(* IEC 61131-3 sources: SRCI_CLIENT_PLC/RobotLibrary/Library/POUs/Read/MC_ReadRobotData/Structures, 4 files *)

(* ---- ReadRobotDataOutCmd.st ---- *)
{attribute 'pack_mode' := '1'}
// -------------------------------------------------------------------------
//  SRCI Robot Library
// -------------------------------------------------------------------------
//
//  Object:      ReadRealsOutCmd
//  Author:      Thorsten Brach
//  Date:        2024-08-09
//
//  Description:
//
//
//  Copyright:
//    (C) 2024 Thorsten Brach. All rights reserved
//             Licensed under the MIT License.
//
//  Disclaimer:
//    This project is provided without any guarantee and can be used for
//    private and commercial purposes. Any use is at the user’s
//    own risk and responsibility.
//
// -------------------------------------------------------------------------
TYPE ReadRobotDataOutCmd :
STRUCT
  /// RC manufacturer name
  RCManufacturer       : STRING(20);
  /// RC part number
  RCOrderID            : STRING(20);
  /// RC serial number
  RCSerialNumber       : STRING(16);
  /// RA serial number
  RASerialNumber       : STRING(16);
  /// Robot firmware version in manufacturer -specific format
  RCFirmwareVersion    : STRING(12);
  ///
  /// Version of the server implementation in the format X.X.X (spec table 6-18) (ST-FIX F46: comment missing)
  RCInterpreterVersion : STRING(11); // ST-FIX F163: three numbers 0..255 as text 'M.m.p' (STRING(5) cut two-digit parts)
  /// Version of the SRCI interpreter on the RC as numbers (spec 6.1.2 table 6-11: Major, Minor, Patch) (ST-FIX F163: the text RCInterpreterVersion was decoded from single characters)
  RCInterpreterVersionNumber : VersionStruct;
  /// TRUE = Axis used in Robot FALSE = Axis NOT used. See Table 6-13 for bit assignment
  AxisJointUsed        : AxisJointUsed;
  /// TRUE = Axis used by Robot FALSE = Axis NOT used. See Table 6-13 for bit assignment.
  AxisExternalUsed     : AxisExternalUsed;
  /// TRUE = mm FALSE = ° See Table 6-13 for bit assignment.
  AxisJointUnit        : AxisJointUnit;
  /// TRUE = mm FALSE = ° See Table 6-13 for bit assignment
  AxisExternalUnit     : AxisExternalUnit;
  /// • TRUE: Function is supported by RC • FALSE: Function is not supported by RC See Table 6-14 for bit assignment.
  RCSupportedFunctions  : RCSupportedFunctions;
  /// Unique and unmodifiable identification of the RA.
  RobotID              : STRING(16);
  /// Interpreter task cycle time of the RC [ms]
  InterpreterCycleTime : UINT;
END_STRUCT
END_TYPE

(* ---- ReadRobotDataParCmd.st ---- *)
{attribute 'pack_mode' := '1'}
// -------------------------------------------------------------------------
//  SRCI Robot Library
// -------------------------------------------------------------------------
//
//  Object:      ReadRealsParCmd
//  Author:      Thorsten Brach
//  Date:        2024-08-09
//
//  Description:
//
//
//  Copyright:
//    (C) 2024 Thorsten Brach. All rights reserved
//             Licensed under the MIT License.
//
//  Disclaimer:
//    This project is provided without any guarantee and can be used for
//    private and commercial purposes. Any use is at the user’s
//    own risk and responsibility.
//
// -------------------------------------------------------------------------
TYPE ReadRobotDataParCmd :
STRUCT
END_STRUCT
END_TYPE

(* ---- ReadRobotDataRecvData.st ---- *)
{attribute 'pack_mode' := '1'}
// -------------------------------------------------------------------------
//  SRCI Robot Library
// -------------------------------------------------------------------------
//
//  Object:      ReadRealsRecvData
//  Author:      Thorsten Brach
//  Date:        2024-08-09
//
//  Description:
//
//
//  Copyright:
//    (C) 2024 Thorsten Brach. All rights reserved
//             Licensed under the MIT License.
//
//  Disclaimer:
//    This project is provided without any guarantee and can be used for
//    private and commercial purposes. Any use is at the user’s
//    own risk and responsibility.
//
// -------------------------------------------------------------------------
TYPE ReadRobotDataRecvData EXTENDS RspHeader :
STRUCT
  /// RC manufacturer name
  RCManufacturer       : STRING(20);
  /// RC part number
  RCOrderID            : STRING(20);
  /// RC serial number
  RCSerialNumber       : STRING(16);
  /// RA serial number
  RASerialNumber       : STRING(16);
  /// Robot firmware version in manufacturer -specific format
  RCFirmwareVersion    : STRING(12);
  ///
  RCInterpreterVersion : STRING(11); // ST-FIX F163: three numbers 0..255 as text 'M.m.p' (STRING(5) cut two-digit parts)
  /// Version of the SRCI interpreter on the RC as numbers (spec 6.1.2 table 6-11: Major, Minor, Patch) (ST-FIX F163: the text RCInterpreterVersion was decoded from single characters)
  RCInterpreterVersionNumber : VersionStruct;
  /// Reserve
  Reserve              : BYTE;
  /// TRUE = Axis used in Robot FALSE = Axis NOT used. See Table 6-13 for bit assignment
  AxisJointUsed        : BYTE;
  /// TRUE = Axis used by Robot FALSE = Axis NOT used. See Table 6-13 for bit assignment.
  AxisExternalUsed     : BYTE;
  /// TRUE = mm FALSE = ° See Table 6-13 for bit assignment.
  AxisJointUnit        : BYTE;
  /// TRUE = mm FALSE = ° See Table 6-13 for bit assignment
  AxisExternalUnit     : BYTE;
  /// • TRUE: Function is supported by RC • FALSE: Function is not supported by RC See Table 6-14 for bit assignment.
  RCSupportedFunctions : ARRAY[0..18] OF BYTE;
  /// Reserve 2
  Reserve2             : BYTE;
  /// Unique and unmodifiable identification of the RA.
  RobotID              : STRING(16);
  /// Interpreter task cycle time of the RC [ms]
  InterpreterCycleTime : UINT;
END_STRUCT
END_TYPE

(* ---- ReadRobotDataSendData.st ---- *)
{attribute 'pack_mode' := '1'}
// -------------------------------------------------------------------------
//  SRCI Robot Library
// -------------------------------------------------------------------------
//
//  Object:      ReadRealsSendData
//  Author:      Thorsten Brach
//  Date:        2024-08-09
//
//  Description:
//
//
//  Copyright:
//    (C) 2024 Thorsten Brach. All rights reserved
//             Licensed under the MIT License.
//
//  Disclaimer:
//    This project is provided without any guarantee and can be used for
//    private and commercial purposes. Any use is at the user’s
//    own risk and responsibility.
//
// -------------------------------------------------------------------------
TYPE ReadRobotDataSendData EXTENDS CmdHeader:
STRUCT
END_STRUCT
END_TYPE
